FUNCTION_BLOCK PID_MODEL_TUNER (* Experimental; offline checks only; native export/runtime pending *)
  (* Standard: 61499-2 *)
  (* Version 0.1, 2026-10-20, Guilherme *)
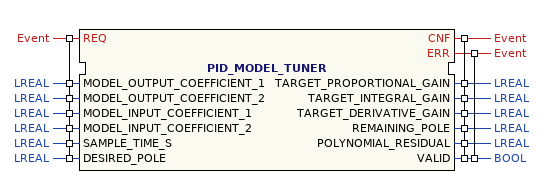
  EVENT_INPUT
    REQ WITH MODEL_OUTPUT_COEFFICIENT_1, MODEL_OUTPUT_COEFFICIENT_2, MODEL_INPUT_COEFFICIENT_1, MODEL_INPUT_COEFFICIENT_2, SAMPLE_TIME_S, DESIRED_POLE;
  END_EVENT
  EVENT_OUTPUT
    CNF WITH TARGET_PROPORTIONAL_GAIN, TARGET_INTEGRAL_GAIN, TARGET_DERIVATIVE_GAIN, REMAINING_POLE, POLYNOMIAL_RESIDUAL, VALID;
    ERR WITH VALID;
  END_EVENT
  VAR_INPUT
    MODEL_OUTPUT_COEFFICIENT_1 : LREAL;
    MODEL_OUTPUT_COEFFICIENT_2 : LREAL;
    MODEL_INPUT_COEFFICIENT_1 : LREAL;
    MODEL_INPUT_COEFFICIENT_2 : LREAL;
    SAMPLE_TIME_S : LREAL;
    DESIRED_POLE : LREAL;
  END_VAR
  VAR_OUTPUT
    TARGET_PROPORTIONAL_GAIN : LREAL;
    TARGET_INTEGRAL_GAIN : LREAL;
    TARGET_DERIVATIVE_GAIN : LREAL;
    REMAINING_POLE : LREAL;
    POLYNOMIAL_RESIDUAL : LREAL;
    VALID : BOOL;
  END_VAR
  VAR
    A1 : LREAL;
    A2 : LREAL;
    B1 : LREAL;
    B2 : LREAL;
    P : LREAL;
    C1 : LREAL;
    C2 : LREAL;
    C3 : LREAL;
    H0 : LREAL;
    H1 : LREAL;
    H2 : LREAL;
    H3 : LREAL;
    S0 : LREAL;
    S1 : LREAL;
    S2 : LREAL;
    T0 : LREAL;
    T1 : LREAL;
    T2 : LREAL;
    DEN : LREAL;
    SCALE : LREAL;
    Q0 : LREAL;
    Q1 : LREAL;
    Q2 : LREAL;
    R : LREAL;
    KP : LREAL;
    KI : LREAL;
    KD : LREAL;
    RES : LREAL;
    MAG : LREAL;
    V1 : LREAL;
    V2 : LREAL;
    V3 : LREAL;
    V4 : LREAL;
  END_VAR
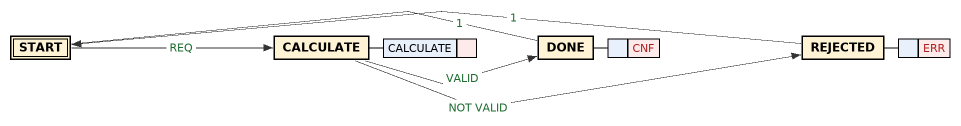
  EC_STATES
    START;
    CALCULATE : CALCULATE;
    DONE : -> CNF;
    REJECTED : -> ERR;
  END_STATES
  EC_TRANSITIONS
    START TO CALCULATE := REQ;
    CALCULATE TO DONE := VALID;
    CALCULATE TO REJECTED := NOT VALID;
    DONE TO START := 1;
    REJECTED TO START := 1;
  END_TRANSITIONS
  ALGORITHM CALCULATE IN ST:
VALID := (MODEL_OUTPUT_COEFFICIENT_1 >= -1.0E+100) AND (MODEL_OUTPUT_COEFFICIENT_1 <= 1.0E+100) AND (MODEL_OUTPUT_COEFFICIENT_2 >= -1.0E+100) AND (MODEL_OUTPUT_COEFFICIENT_2 <= 1.0E+100) AND (MODEL_INPUT_COEFFICIENT_1 >= -1.0E+100) AND (MODEL_INPUT_COEFFICIENT_1 <= 1.0E+100) AND (MODEL_INPUT_COEFFICIENT_2 >= -1.0E+100) AND (MODEL_INPUT_COEFFICIENT_2 <= 1.0E+100) AND (SAMPLE_TIME_S >= -1.0E+100) AND (SAMPLE_TIME_S <= 1.0E+100) AND (DESIRED_POLE >= -1.0E+100) AND (DESIRED_POLE <= 1.0E+100) AND (SAMPLE_TIME_S > 0.0) AND (DESIRED_POLE > 0.0) AND (DESIRED_POLE < 1.0);
IF VALID THEN
A1 := MODEL_OUTPUT_COEFFICIENT_1;
A2 := MODEL_OUTPUT_COEFFICIENT_2;
B1 := MODEL_INPUT_COEFFICIENT_1;
B2 := MODEL_INPUT_COEFFICIENT_2;
P := DESIRED_POLE;
SCALE := B1;
IF SCALE < 0.0 THEN
SCALE := -SCALE;
END_IF;
MAG := B2;
IF MAG < 0.0 THEN
MAG := -MAG;
END_IF;
IF MAG > SCALE THEN
SCALE := MAG;
END_IF;
MAG := B1;
IF MAG < 0.0 THEN
MAG := -MAG;
END_IF;
VALID := (SCALE > 1.0E-12) AND (MAG > 1.0E-10 * SCALE);
IF VALID THEN
C1 := -3.0 * P;
C2 := 3.0 * P * P;
C3 := -P * P * P;
H0 := C1 + 1.0 + A1;
H1 := C2 - A1 + A2;
H2 := C3 - A2;
H3 := 0.0;
S0 := H0 / B1;
T0 := -1.0 / B1;
S1 := (H1 - B2 * S0) / B1;
T1 := (-C1 - B2 * T0) / B1;
S2 := (H2 - B2 * S1) / B1;
T2 := (-C2 - B2 * T1) / B1;
DEN := B2 * T2 + C3;
SCALE := B2 * T2;
IF SCALE < 0.0 THEN
SCALE := -SCALE;
END_IF;
MAG := C3;
IF MAG < 0.0 THEN
MAG := -MAG;
END_IF;
SCALE := SCALE + MAG;
MAG := DEN;
IF MAG < 0.0 THEN
MAG := -MAG;
END_IF;
VALID := (S0 >= -1.0E+100) AND (S0 <= 1.0E+100) AND (S1 >= -1.0E+100) AND (S1 <= 1.0E+100) AND (S2 >= -1.0E+100) AND (S2 <= 1.0E+100) AND (T0 >= -1.0E+100) AND (T0 <= 1.0E+100) AND (T1 >= -1.0E+100) AND (T1 <= 1.0E+100) AND (T2 >= -1.0E+100) AND (T2 <= 1.0E+100) AND (DEN >= -1.0E+100) AND (DEN <= 1.0E+100) AND (SCALE >= -1.0E+100) AND (SCALE <= 1.0E+100) AND (MAG > 1.0E-10 * SCALE) AND (MAG > 1.0E-12);
IF VALID THEN
R := (H3 - B2 * S2) / DEN;
Q0 := S0 + T0 * R;
Q1 := S1 + T1 * R;
Q2 := S2 + T2 * R;
KP := (Q0 - Q1 - 3.0 * Q2) / 2.0;
KI := (Q0 + Q1 + Q2) / SAMPLE_TIME_S;
KD := SAMPLE_TIME_S * Q2;
V1 := -1.0 - A1 + B1 * Q0 - (C1 - R);
V2 := A1 - A2 + B1 * Q1 + B2 * Q0 - (C2 - C1 * R);
V3 := A2 + B1 * Q2 + B2 * Q1 - (C3 - C2 * R);
V4 := B2 * Q2 + C3 * R;
RES := 0.0;
MAG := V1;
IF MAG < 0.0 THEN
MAG := -MAG;
END_IF;
IF MAG > RES THEN
RES := MAG;
END_IF;
MAG := V2;
IF MAG < 0.0 THEN
MAG := -MAG;
END_IF;
IF MAG > RES THEN
RES := MAG;
END_IF;
MAG := V3;
IF MAG < 0.0 THEN
MAG := -MAG;
END_IF;
IF MAG > RES THEN
RES := MAG;
END_IF;
MAG := V4;
IF MAG < 0.0 THEN
MAG := -MAG;
END_IF;
IF MAG > RES THEN
RES := MAG;
END_IF;
VALID := (R >= -1.0E+100) AND (R <= 1.0E+100) AND (Q0 >= -1.0E+100) AND (Q0 <= 1.0E+100) AND (Q1 >= -1.0E+100) AND (Q1 <= 1.0E+100) AND (Q2 >= -1.0E+100) AND (Q2 <= 1.0E+100) AND (KP >= -1.0E+100) AND (KP <= 1.0E+100) AND (KI >= -1.0E+100) AND (KI <= 1.0E+100) AND (KD >= -1.0E+100) AND (KD <= 1.0E+100) AND (V1 >= -1.0E+100) AND (V1 <= 1.0E+100) AND (V2 >= -1.0E+100) AND (V2 <= 1.0E+100) AND (V3 >= -1.0E+100) AND (V3 <= 1.0E+100) AND (V4 >= -1.0E+100) AND (V4 <= 1.0E+100) AND (RES >= -1.0E+100) AND (RES <= 1.0E+100) AND (R > -1.0) AND (R < 1.0) AND (KP >= 0.0) AND (KI >= 0.0) AND (KD >= 0.0) AND (RES <= 1.0E-9);
IF VALID THEN
TARGET_PROPORTIONAL_GAIN := KP;
TARGET_INTEGRAL_GAIN := KI;
TARGET_DERIVATIVE_GAIN := KD;
REMAINING_POLE := R;
POLYNOMIAL_RESIDUAL := RES;
END_IF;
END_IF;
END_IF;
END_IF;
  END_ALGORITHM
END_FUNCTION_BLOCK
